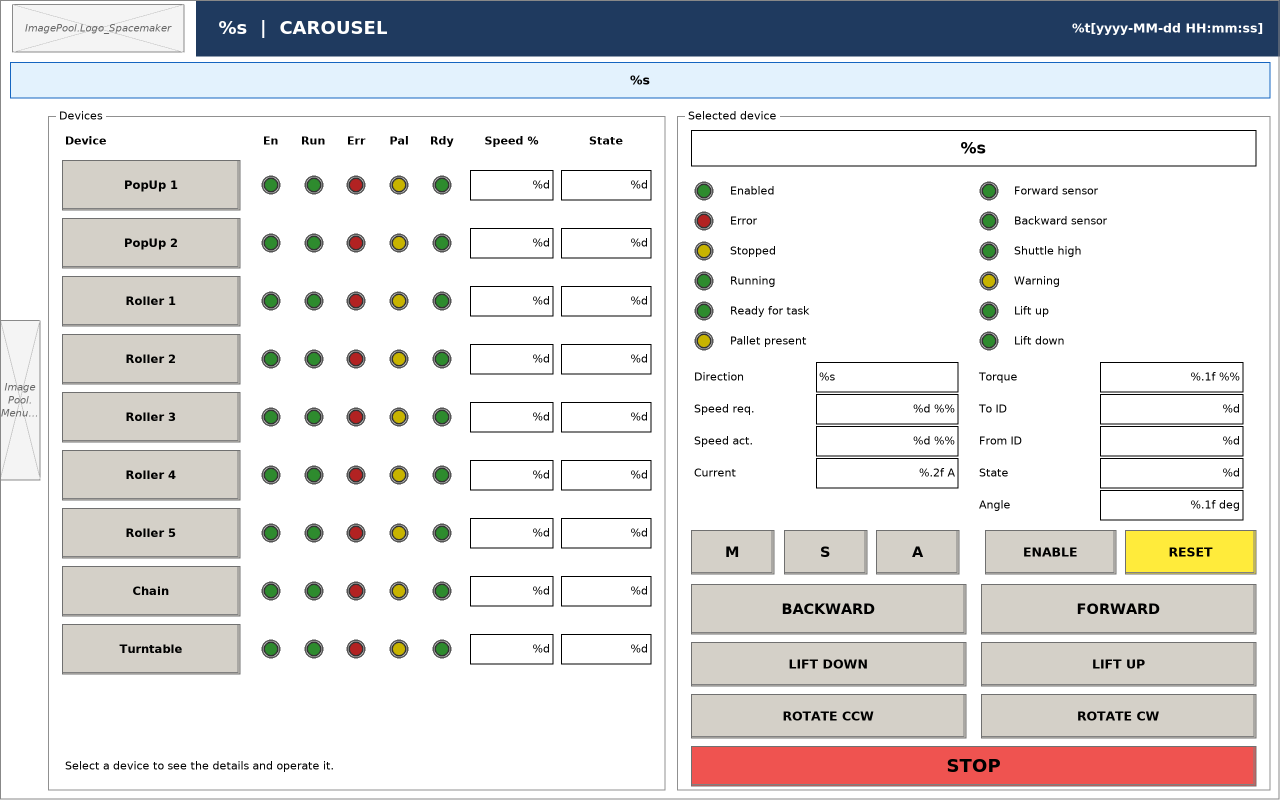
VISUALIZATION Carrousel  // 1280x800
    Rectangle (0,0 196x56)
        OnMouseClick: change screen: Main
    Image (12,4 172x48), image: ImagePool.Logo_Spacemaker
        OnMouseClick: change screen: Main
    Rectangle (196,0 1084x56), "%s | CAROUSEL", text variable: GVL_HMI_System.stStatus.sSystemName
    Rectangle (930,8 336x40), "%t[yyyy-MM-dd HH:mm:ss]", text variable: GVL_HMI_System.stStatus.dtNow
    Rectangle (10,62 1260x36), "%s", text variable: GVL_HMI_System.stStatus.sMessage, colour toggle: GVL_HMI_System.stStatus.bMessageAlarm
    GroupBox (48,108 617x682), "Devices"
    Rectangle (62,128 178x26), "Device"
    Rectangle (250,128 42x26), "En"
    Rectangle (292,128 43x26), "Run"
    Rectangle (335,128 43x26), "Err"
    Rectangle (378,128 43x26), "Pal"
    Rectangle (421,128 42x26), "Rdy"
    Rectangle (470,128 83x26), "Speed %"
    Rectangle (561,128 90x26), "State"
    Button (62,160 178x50), "PopUp 1", colour toggle: GVL_HMI_Carousel.astDevice[1].bSelected
        OnMouseClick: execute { GVL_HMI_Carousel.uiSelected := 1; }
    Lamp1 (260,174 22x22), variable: GVL_HMI_Carousel.astDevice[1].bEnabled, style: Lamp-Lamp1-Green
    Lamp1 (303,174 22x22), variable: GVL_HMI_Carousel.astDevice[1].bRunning, style: Lamp-Lamp1-Green
    Lamp1 (345,174 22x22), variable: GVL_HMI_Carousel.astDevice[1].bError, style: Lamp-Lamp1-Red
    Lamp1 (388,174 22x22), variable: GVL_HMI_Carousel.astDevice[1].bOccupied, style: Lamp-Lamp1-Yellow
    Lamp1 (431,174 22x22), variable: GVL_HMI_Carousel.astDevice[1].bReadyForTask, style: Lamp-Lamp1-Green
    Rectangle (470,170 83x30), "%d", text variable: GVL_HMI_Carousel.astDevice[1].iSpeedActual_pct
    Rectangle (561,170 90x30), "%d", text variable: GVL_HMI_Carousel.astDevice[1].uiStateMachine
    Button (62,218 178x50), "PopUp 2", colour toggle: GVL_HMI_Carousel.astDevice[2].bSelected
        OnMouseClick: execute { GVL_HMI_Carousel.uiSelected := 2; }
    Lamp1 (260,232 22x22), variable: GVL_HMI_Carousel.astDevice[2].bEnabled, style: Lamp-Lamp1-Green
    Lamp1 (303,232 22x22), variable: GVL_HMI_Carousel.astDevice[2].bRunning, style: Lamp-Lamp1-Green
    Lamp1 (345,232 22x22), variable: GVL_HMI_Carousel.astDevice[2].bError, style: Lamp-Lamp1-Red
    Lamp1 (388,232 22x22), variable: GVL_HMI_Carousel.astDevice[2].bOccupied, style: Lamp-Lamp1-Yellow
    Lamp1 (431,232 22x22), variable: GVL_HMI_Carousel.astDevice[2].bReadyForTask, style: Lamp-Lamp1-Green
    Rectangle (470,228 83x30), "%d", text variable: GVL_HMI_Carousel.astDevice[2].iSpeedActual_pct
    Rectangle (561,228 90x30), "%d", text variable: GVL_HMI_Carousel.astDevice[2].uiStateMachine
    Button (62,276 178x50), "Roller 1", colour toggle: GVL_HMI_Carousel.astDevice[3].bSelected
        OnMouseClick: execute { GVL_HMI_Carousel.uiSelected := 3; }
    Lamp1 (260,290 22x22), variable: GVL_HMI_Carousel.astDevice[3].bEnabled, style: Lamp-Lamp1-Green
    Lamp1 (303,290 22x22), variable: GVL_HMI_Carousel.astDevice[3].bRunning, style: Lamp-Lamp1-Green
    Lamp1 (345,290 22x22), variable: GVL_HMI_Carousel.astDevice[3].bError, style: Lamp-Lamp1-Red
    Lamp1 (388,290 22x22), variable: GVL_HMI_Carousel.astDevice[3].bOccupied, style: Lamp-Lamp1-Yellow
    Lamp1 (431,290 22x22), variable: GVL_HMI_Carousel.astDevice[3].bReadyForTask, style: Lamp-Lamp1-Green
    Rectangle (470,286 83x30), "%d", text variable: GVL_HMI_Carousel.astDevice[3].iSpeedActual_pct
    Rectangle (561,286 90x30), "%d", text variable: GVL_HMI_Carousel.astDevice[3].uiStateMachine
    Button (62,334 178x50), "Roller 2", colour toggle: GVL_HMI_Carousel.astDevice[4].bSelected
        OnMouseClick: execute { GVL_HMI_Carousel.uiSelected := 4; }
    Lamp1 (260,348 22x22), variable: GVL_HMI_Carousel.astDevice[4].bEnabled, style: Lamp-Lamp1-Green
    Lamp1 (303,348 22x22), variable: GVL_HMI_Carousel.astDevice[4].bRunning, style: Lamp-Lamp1-Green
    Lamp1 (345,348 22x22), variable: GVL_HMI_Carousel.astDevice[4].bError, style: Lamp-Lamp1-Red
    Lamp1 (388,348 22x22), variable: GVL_HMI_Carousel.astDevice[4].bOccupied, style: Lamp-Lamp1-Yellow
    Lamp1 (431,348 22x22), variable: GVL_HMI_Carousel.astDevice[4].bReadyForTask, style: Lamp-Lamp1-Green
    Rectangle (470,344 83x30), "%d", text variable: GVL_HMI_Carousel.astDevice[4].iSpeedActual_pct
    Rectangle (561,344 90x30), "%d", text variable: GVL_HMI_Carousel.astDevice[4].uiStateMachine
    Button (62,392 178x50), "Roller 3", colour toggle: GVL_HMI_Carousel.astDevice[5].bSelected
        OnMouseClick: execute { GVL_HMI_Carousel.uiSelected := 5; }
    Lamp1 (260,406 22x22), variable: GVL_HMI_Carousel.astDevice[5].bEnabled, style: Lamp-Lamp1-Green
    Lamp1 (303,406 22x22), variable: GVL_HMI_Carousel.astDevice[5].bRunning, style: Lamp-Lamp1-Green
    Lamp1 (345,406 22x22), variable: GVL_HMI_Carousel.astDevice[5].bError, style: Lamp-Lamp1-Red
    Lamp1 (388,406 22x22), variable: GVL_HMI_Carousel.astDevice[5].bOccupied, style: Lamp-Lamp1-Yellow
    Lamp1 (431,406 22x22), variable: GVL_HMI_Carousel.astDevice[5].bReadyForTask, style: Lamp-Lamp1-Green
    Rectangle (470,402 83x30), "%d", text variable: GVL_HMI_Carousel.astDevice[5].iSpeedActual_pct
    Rectangle (561,402 90x30), "%d", text variable: GVL_HMI_Carousel.astDevice[5].uiStateMachine
    Button (62,450 178x50), "Roller 4", colour toggle: GVL_HMI_Carousel.astDevice[6].bSelected
        OnMouseClick: execute { GVL_HMI_Carousel.uiSelected := 6; }
    Lamp1 (260,464 22x22), variable: GVL_HMI_Carousel.astDevice[6].bEnabled, style: Lamp-Lamp1-Green
    Lamp1 (303,464 22x22), variable: GVL_HMI_Carousel.astDevice[6].bRunning, style: Lamp-Lamp1-Green
    Lamp1 (345,464 22x22), variable: GVL_HMI_Carousel.astDevice[6].bError, style: Lamp-Lamp1-Red
    Lamp1 (388,464 22x22), variable: GVL_HMI_Carousel.astDevice[6].bOccupied, style: Lamp-Lamp1-Yellow
    Lamp1 (431,464 22x22), variable: GVL_HMI_Carousel.astDevice[6].bReadyForTask, style: Lamp-Lamp1-Green
    Rectangle (470,460 83x30), "%d", text variable: GVL_HMI_Carousel.astDevice[6].iSpeedActual_pct
    Rectangle (561,460 90x30), "%d", text variable: GVL_HMI_Carousel.astDevice[6].uiStateMachine
    Button (62,508 178x50), "Roller 5", colour toggle: GVL_HMI_Carousel.astDevice[7].bSelected
        OnMouseClick: execute { GVL_HMI_Carousel.uiSelected := 7; }
    Lamp1 (260,522 22x22), variable: GVL_HMI_Carousel.astDevice[7].bEnabled, style: Lamp-Lamp1-Green
    Lamp1 (303,522 22x22), variable: GVL_HMI_Carousel.astDevice[7].bRunning, style: Lamp-Lamp1-Green
    Lamp1 (345,522 22x22), variable: GVL_HMI_Carousel.astDevice[7].bError, style: Lamp-Lamp1-Red
    Lamp1 (388,522 22x22), variable: GVL_HMI_Carousel.astDevice[7].bOccupied, style: Lamp-Lamp1-Yellow
    Lamp1 (431,522 22x22), variable: GVL_HMI_Carousel.astDevice[7].bReadyForTask, style: Lamp-Lamp1-Green
    Rectangle (470,518 83x30), "%d", text variable: GVL_HMI_Carousel.astDevice[7].iSpeedActual_pct
    Rectangle (561,518 90x30), "%d", text variable: GVL_HMI_Carousel.astDevice[7].uiStateMachine
    Button (62,566 178x50), "Chain", colour toggle: GVL_HMI_Carousel.astDevice[8].bSelected
        OnMouseClick: execute { GVL_HMI_Carousel.uiSelected := 8; }
    Lamp1 (260,580 22x22), variable: GVL_HMI_Carousel.astDevice[8].bEnabled, style: Lamp-Lamp1-Green
    Lamp1 (303,580 22x22), variable: GVL_HMI_Carousel.astDevice[8].bRunning, style: Lamp-Lamp1-Green
    Lamp1 (345,580 22x22), variable: GVL_HMI_Carousel.astDevice[8].bError, style: Lamp-Lamp1-Red
    Lamp1 (388,580 22x22), variable: GVL_HMI_Carousel.astDevice[8].bOccupied, style: Lamp-Lamp1-Yellow
    Lamp1 (431,580 22x22), variable: GVL_HMI_Carousel.astDevice[8].bReadyForTask, style: Lamp-Lamp1-Green
    Rectangle (470,576 83x30), "%d", text variable: GVL_HMI_Carousel.astDevice[8].iSpeedActual_pct
    Rectangle (561,576 90x30), "%d", text variable: GVL_HMI_Carousel.astDevice[8].uiStateMachine
    Button (62,624 178x50), "Turntable", colour toggle: GVL_HMI_Carousel.astDevice[9].bSelected
        OnMouseClick: execute { GVL_HMI_Carousel.uiSelected := 9; }
    Lamp1 (260,638 22x22), variable: GVL_HMI_Carousel.astDevice[9].bEnabled, style: Lamp-Lamp1-Green
    Lamp1 (303,638 22x22), variable: GVL_HMI_Carousel.astDevice[9].bRunning, style: Lamp-Lamp1-Green
    Lamp1 (345,638 22x22), variable: GVL_HMI_Carousel.astDevice[9].bError, style: Lamp-Lamp1-Red
    Lamp1 (388,638 22x22), variable: GVL_HMI_Carousel.astDevice[9].bOccupied, style: Lamp-Lamp1-Yellow
    Lamp1 (431,638 22x22), variable: GVL_HMI_Carousel.astDevice[9].bReadyForTask, style: Lamp-Lamp1-Green
    Rectangle (470,634 83x30), "%d", text variable: GVL_HMI_Carousel.astDevice[9].iSpeedActual_pct
    Rectangle (561,634 90x30), "%d", text variable: GVL_HMI_Carousel.astDevice[9].uiStateMachine
    Rectangle (62,752 593x28), "Select a device to see the details and operate it."
    GroupBox (677,108 593x682), "Selected device"
    Rectangle (691,130 565x36), "%s", text variable: GVL_HMI_Carousel.stSelected.sName
    Lamp1 (693,180 22x22), variable: GVL_HMI_Carousel.stSelected.bEnabled, style: Lamp-Lamp1-Green
    Rectangle (727,176 201x30), "Enabled"
    Lamp1 (693,210 22x22), variable: GVL_HMI_Carousel.stSelected.bError, style: Lamp-Lamp1-Red
    Rectangle (727,206 201x30), "Error"
    Lamp1 (693,240 22x22), variable: GVL_HMI_Carousel.stSelected.bStopped, style: Lamp-Lamp1-Yellow
    Rectangle (727,236 201x30), "Stopped"
    Lamp1 (693,270 22x22), variable: GVL_HMI_Carousel.stSelected.bRunning, style: Lamp-Lamp1-Green
    Rectangle (727,266 201x30), "Running"
    Lamp1 (693,300 22x22), variable: GVL_HMI_Carousel.stSelected.bReadyForTask, style: Lamp-Lamp1-Green
    Rectangle (727,296 201x30), "Ready for task"
    Lamp1 (693,330 22x22), variable: GVL_HMI_Carousel.stSelected.bOccupied, style: Lamp-Lamp1-Yellow
    Rectangle (727,326 201x30), "Pallet present"
    Lamp1 (978,180 22x22), variable: GVL_HMI_Carousel.stSelected.bForwardSensor, style: Lamp-Lamp1-Green
    Rectangle (1011,176 202x30), "Forward sensor"
    Lamp1 (978,210 22x22), variable: GVL_HMI_Carousel.stSelected.bBackwardSensor, style: Lamp-Lamp1-Green
    Rectangle (1011,206 202x30), "Backward sensor"
    Lamp1 (978,240 22x22), variable: GVL_HMI_Carousel.stSelected.bShuttleHigh, style: Lamp-Lamp1-Green
    Rectangle (1011,236 202x30), "Shuttle high"
    Lamp1 (978,270 22x22), variable: GVL_HMI_Carousel.stSelected.bWarning, style: Lamp-Lamp1-Yellow
    Rectangle (1011,266 202x30), "Warning"
    Lamp1 (978,300 22x22), variable: GVL_HMI_Carousel.stSelected.bLiftUp, style: Lamp-Lamp1-Green
    Rectangle (1011,296 202x30), "Lift up"
    Lamp1 (978,330 22x22), variable: GVL_HMI_Carousel.stSelected.bLiftDown, style: Lamp-Lamp1-Green
    Rectangle (1011,326 202x30), "Lift down"
    Rectangle (691,362 119x30), "Direction"
    Rectangle (816,362 142x30), "%s", text variable: GVL_HMI_Carousel.stSelected.sMotorDirection
    Rectangle (691,394 119x30), "Speed req."
    Rectangle (816,394 142x30), "%d %%", text variable: GVL_HMI_Carousel.stSelected.iSpeedRequested_pct
    Rectangle (691,426 119x30), "Speed act."
    Rectangle (816,426 142x30), "%d %%", text variable: GVL_HMI_Carousel.stSelected.iSpeedActual_pct
    Rectangle (691,458 119x30), "Current"
    Rectangle (816,458 142x30), "%.2f A", text variable: GVL_HMI_Carousel.stSelected.rCurrent_A
    Rectangle (976,362 118x30), "Torque"
    Rectangle (1100,362 143x30), "%.1f %%", text variable: GVL_HMI_Carousel.stSelected.rTorque_pct
    Rectangle (976,394 118x30), "To ID"
    Rectangle (1100,394 143x30), "%d", text variable: GVL_HMI_Carousel.stSelected.diTransferToId
    Rectangle (976,426 118x30), "From ID"
    Rectangle (1100,426 143x30), "%d", text variable: GVL_HMI_Carousel.stSelected.diTransferFromId
    Rectangle (976,458 118x30), "State"
    Rectangle (1100,458 143x30), "%d", text variable: GVL_HMI_Carousel.stSelected.uiStateMachine
    Rectangle (976,490 118x30), "Angle"
    Rectangle (1100,490 143x30), "%.1f deg", text variable: GVL_HMI_Carousel.stSelected.rAngle_deg
    Button (691,530 83x44), "M", colour toggle: GVL_HMI_Carousel.stSelected.bModeManual
        tap GVL_HMI_Carousel.stCommand.bModeManual p3779583253=TRUE
    Button (784,530 83x44), "S", colour toggle: GVL_HMI_Carousel.stSelected.bModeSemi
        tap GVL_HMI_Carousel.stCommand.bModeSemi p3779583253=TRUE
    Button (876,530 83x44), "A", colour toggle: GVL_HMI_Carousel.stSelected.bModeAuto
        tap GVL_HMI_Carousel.stCommand.bModeAuto p3779583253=TRUE
    Button (985,530 131x44), "ENABLE", colour toggle: GVL_HMI_Carousel.stSelected.bEnabled
        tap GVL_HMI_Carousel.stCommand.bEnable p3779583253=TRUE
    Button (1125,530 131x44), "RESET"
        tap GVL_HMI_Carousel.stCommand.bReset p3779583253=TRUE
    Button (691,584 275x50), "BACKWARD", input disabled if: NOT GVL_HMI_Carousel.stSelected.bModeManual
        tap GVL_HMI_Carousel.stCommand.bJogBackward p3779583253=TRUE
    Button (981,584 275x50), "FORWARD", input disabled if: NOT GVL_HMI_Carousel.stSelected.bModeManual
        tap GVL_HMI_Carousel.stCommand.bJogForward p3779583253=TRUE
    Button (691,642 275x44), "LIFT DOWN", input disabled if: NOT GVL_HMI_Carousel.stSelected.bHasLift
        tap GVL_HMI_Carousel.stCommand.bLiftDown p3779583253=TRUE
    Button (981,642 275x44), "LIFT UP", input disabled if: NOT GVL_HMI_Carousel.stSelected.bHasLift
        tap GVL_HMI_Carousel.stCommand.bLiftUp p3779583253=TRUE
    Button (691,694 275x44), "ROTATE CCW", input disabled if: NOT GVL_HMI_Carousel.stSelected.bHasRotation
        tap GVL_HMI_Carousel.stCommand.bRotateCcw p3779583253=TRUE
    Button (981,694 275x44), "ROTATE CW", input disabled if: NOT GVL_HMI_Carousel.stSelected.bHasRotation
        tap GVL_HMI_Carousel.stCommand.bRotateCw p3779583253=TRUE
    Button (691,746 565x40), "STOP"
        tap GVL_HMI_Carousel.stCommand.bStop p3779583253=TRUE
    Rectangle (0,320 40x160)
        OnMouseEnter: OpenDialog Dialog=Dialog, OpenModal=True, PositionX=0, PositionY=0
        OnMouseClick: OpenDialog Dialog=Dialog, OpenModal=True, PositionX=0, PositionY=0
    Image (0,320 40x160), image: ImagePool.Menu_Tab
        OnMouseEnter: OpenDialog Dialog=Dialog, OpenModal=True, PositionX=0, PositionY=0
        OnMouseClick: OpenDialog Dialog=Dialog, OpenModal=True, PositionX=0, PositionY=0
END_VISUALIZATION

(* stored: Version 1.1.0.1
   Visu Carrousel: Id {c5170854-078b-4555-90ff-62533ca7440d} *)
